Fanuc KAREL source: KT00400.KL

PROGRAM KT00400
%NOLOCKGROUP
VAR
  C1: CONFIG
  C2: CONFIG
  OUT: BOOLEAN
BEGIN
  C1.CFG_FLIP = TRUE
  C2.CFG_FLIP = FALSE
  C1.CFG_FLIP = TRUE
  C2.CFG_FLIP = FALSE
  OUT = C1 <= C2
END KT00400
